Staubli VAL3: onStart.pgx

program onStart()
  local num l_i
  local string l_sPath
  local num i
begin
  l_sPath="Disk://data/CustomerLib"
  libList(l_sPath,sLibList)

  resize(sList,1,size(savedata:tToolItem))

  bIsDoing=false
  for l_i = 0 to size(sList)-1
    sList[l_i]=toString("",l_i)+","+savedata:tToolItem[l_i].sName
  endFor

  sSelTool=toString("",savedata:nUsingTool)+","+savedata:tToolItem[savedata:nUsingTool].sName
  sLastTool=""
//  bLock=true
//  sBtnUnLock="解锁"
//  //获取机器人类型
//  call libTqe:_getArmType(sArmType,sArmDetail)
//  if sArmType=="4_Axis"
//    resize(bDisable,1,4)
//    resize(nMaxJntForec,1,4)
//    bSix_Axis=false
//  elseIf sArmType=="6_Axis"
//    resize(bDisable,1,6)
//    resize(nMaxJntForec,1,6)
//    bSix_Axis=true
//  endIf
//  //初始化扭矩设置解锁按钮
//  for i=0 to size(bDisable)-1
//    bDisable[i]=true
//  endFor
  //  call libTqe:_getSetForce(nMaxJntForec)
  call libTqe:initParameter()
end
